// TIA Portal V17 export
DATA_BLOCK "MCP_RC_DB6"   // DB9806
{ S7_Optimized_Access := 'TRUE' }
   VAR
      Count : Int := 3;
      Bad : "MCP_RC_NoSuchUDT";
   END_VAR
BEGIN
END_DATA_BLOCK
